(* PLC project Vn_literals, Beckhoff Automation GmbH TwinCAT PLC Control 3.5.13.21 *)
(* stored: creationDateTime 1970-01-01T00:00:00 *)

PROGRAM Vn_literals

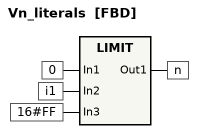
(* FBD diagram, written out as Structured Text *)
n := LIMIT(0, i1, 16#FF);
END_PROGRAM
